Fanuc KAREL source: KA00208.KL

PROGRAM KA00208
%NOLOCKGROUP
VAR
  SRC: ARRAY[4] OF XYZWPR
  DST: ARRAY[4] OF INTEGER
BEGIN
  DST = SRC
END KA00208
